FUNCTION_BLOCK FB_DomeParkingState EXTENDS FB_DomeState

VAR
	Stage		: UINT:= 0;
	tonTimeout	: TON:= (PT:=T#3M); // see Baader Handbook
	tonSleep	: TON := (PT:=T#2S);
	tonDelay	: TON:= (PT:=T#20MS);
	
	sSeperator		: STRING := 'd#azi';
	sLeft			: STRING;
	sAzi			: STRING;
	fAzi			: LREAL;
	fAzi_Old		: LREAL;
	bSplitSuccess 	: BOOL;
END_VAR


METHOD CloseCommand : BOOL
Stage := 0;
tonSleep(IN:=FALSE);
tonTimeout(IN:=FALSE);
tonDelay(IN:=FALSE);
pDome^.SetState(pDome^.fbDomeCloseingState);
END_METHOD


METHOD FoundError : BOOL
Stage:= 0;
tonSleep(IN:=FALSE);
tonTimeout(IN:=FALSE);
tonDelay(IN:=FALSE);
pDome^._Error := TRUE;
pDome^.SetState(pDome^.fbDomeErrorState);
END_METHOD

METHOD OpenCommand : BOOL
Stage:= 0;
tonSleep(IN:=FALSE);
tonTimeout(IN:=FALSE);
tonDelay(IN:=FALSE);
pDome^.SetState(pDome^.fbDomeOpeningState);
END_METHOD

METHOD RunState : BOOL
VAR_INPUT
END_VAR
CASE Stage OF
	0:
		tonTimeout(IN:=TRUE);
		IF NOT pDome^.fbReceive.Busy AND NOT pDome^.fbSend.Busy THEN
			Stage := 1;
		END_IF
	1:
		pDome^.fbSend(	SendString:= 'd#azi0000',
					TXbuffer:= TxBufferDome,
					Busy=>,
					Error=> );
		IF NOT pDome^.fbSend.Busy  THEN
			Stage := 2;
		END_IF
	2:
		IF pDome^._HasReceivedString THEN
			IF pDome^._ReceivedString = 'd#comerro' OR pDome^._ReceivedString = 'd#domerro' THEN
				FoundError();
			ELSIF pDome^._ReceivedString = 'd#gotmess' THEN
				Stage := 3;
			END_IF
		ELSIF NOT pDome^.fbReceive.Busy THEN
			tonSleep(IN:=TRUE);
			IF tonSleep.Q THEN
				tonSleep(IN:=FALSE);
				Stage := 1;
			END_IF
		END_IF
		tonTimeout(IN:=TRUE);
		IF tonTimeout.Q THEN
			tonTimeout(IN:=FALSE);
			FoundError();
		END_IF
	3:
		tonTimeout(IN:=FALSE);
		tonSleep(IN:=TRUE);
		IF tonSleep.Q THEN
			tonSleep(IN:=FALSE);
			Stage := 4;
			tonTimeout(IN:=TRUE);
		END_IF
	4:
		pDome^.fbSend(	SendString:= 'd#getazim',
					TXbuffer:= TxBufferDome,
					Busy=>,
					Error=> );
		IF NOT pDome^.fbSend.Busy  THEN
			Stage := 5;
		END_IF
	5: 
		IF pDome^._HasReceivedString THEN
			IF pDome^._ReceivedString = 'd#comerro' OR pDome^._ReceivedString = 'd#domerro' THEN
				FoundError();
			ELSE
				bSplitSuccess := FindAndSplit(
									pSeparator := ADR(sSeperator),
									pSrcString := ADR(pDome^.sReceivedString),
									pLeftString:= ADR(sLeft),
									nLeftSize	:= 1,
									pRightString := ADR(sAzi),
									nRightSize := 5,
									bSearchFromRight:= FALSE);
				IF bSplitSuccess AND ( STRING_TO_LREAL(sAzi) <> 0 OR sAzi = '0000' ) THEN
					// (STRING_TO_LREAL(sAzi) <> 0 OR sAzi := '0000') -> either sAzi actual 0 OR STRING_TO_LREAL error
					fAzi := STRING_TO_LREAL(sAzi)/10.0;
					//Baader measures azimuth as West of South, so we need to convert it. This works both ways.
					IF fAzi  >= 180.0 THEN
						pDome^._Position := fAzi - 180.0;
					ELSE
						pDome^._Position := fAzi + 180.0;
					END_IF
					IF fAzi = fAzi_Old THEN
						IF ABS(pDome^.Position - 180.0) < 5.0 THEN
							pDome^._DomeRotationState := E_DomeRotationState.parked;
							Stage := 6;
						ELSE
							pDome^._DomeRotationState := E_DomeRotationState.idle;
							// stopped but not parked? try again
							Stage := 0;
						END_IF
					ELSE
						pDome^._DomeRotationState := E_DomeRotationState.slewing;
						// carry on
						Stage := 3;
					END_IF
					fAzi_Old := fAzi;
				END_IF
			END_IF
		ELSIF NOT pDome^.fbReceive.Busy THEN
			tonSleep(IN:=TRUE);
			IF tonSleep.Q THEN
				tonSleep(IN:=FALSE);
				Stage := 4;
			END_IF
		END_IF
		tonTimeout(IN:=TRUE);
		IF tonTimeout.Q THEN
			tonTimeout(IN:=FALSE);
			FoundError();
		END_IF
	6:
		tonTimeout(IN:=FALSE);
		SuccessfulFinished();
		
END_CASE
END_METHOD

PROPERTY StateID : STRING
GET
StateID := 'Parking State';
END_GET
END_PROPERTY


METHOD StopCommand : BOOL
Stage:= 0;
tonSleep(IN:=FALSE);
tonTimeout(IN:=FALSE);
tonDelay(IN:=FALSE);
pDome^.SetState(pDome^.fbDomeStoppingState);
END_METHOD


METHOD SuccessfulFinished : BOOL
Stage:= 0;
tonSleep(IN:=FALSE);
tonTimeout(IN:=FALSE);
tonDelay(IN:=FALSE);
pDome^.SetState(pDome^.fbDomeIdleState);
END_METHOD

END_FUNCTION_BLOCK

(* stored: Version 1.1.0.1, ProductVersion 3.1.4024.15
   POU FB_DomeParkingState: Id {38fd3f71-8ee5-411c-9502-503e70ff8fa9}, SpecialFunc None
   Method CloseCommand: Id {6974039e-2ad8-4be3-a7c5-073290f4b5f6}
   Method FoundError: Id {973b9bd2-f8fb-469d-9375-7bbf24d458da}
   Method OpenCommand: Id {9df60541-5e83-447d-86fb-d70ae39cfb87}
   Method RunState: Id {74c4ccf9-d5e0-427f-ae6f-4cf604480af3}
   Property StateID: Id {077ee837-ee21-442d-8c88-4822066bbecc}
   Get Get: Id {06c04b97-ab55-46ea-a2de-63112be1cd2b}
   Method StopCommand: Id {4adfc0bd-0c92-49b3-ad40-a4adba482d47}
   Method SuccessfulFinished: Id {eaa94ad4-58a6-4ca5-9c6f-84da24826579} *)
